(* IEC 61131-3 sources: s7-to-codesys/tests/POUs/ScenariosLang/FB_StarterFbd_ScenarioTest, 10 files *)

(* ---- FB_StarterFbd_ScenarioTest.decl.st ---- *)
// AUTO-GENERATED — не редактировать: s7conv gen-tests, сценарии scenarios/lang/FB_Starter.csv
// Правка — в CSV (scenarios/README.md), затем python -m s7conv build-corpus.
// Назначение: тесты поведения сконвертированного FB_StarterFbd по сценариям CSV (сценариев: 9, строк: 47):
//             один метод-тест на сценарий, строки — по порядку с моделируемым временем GVL_S7Clock.
//             Ожидаемые значения — из CSV (эталонные модели по описанию логики блока), не из
//             результата конвертации.
// Автор:      s7conv 0.1.0 (сгенерировано)
// Версия:     не указана
// Документ:   scenarios/README.md, docs/methodology.md, раздел «Проверка поведения»
FUNCTION_BLOCK FB_StarterFbd_ScenarioTest EXTENDS coUnit.FB_TestSuite
VAR
    fbStartStop : FB_StarterFbd;  // свой экземпляр на сценарий
    xStartStopDone : BOOL;  // сценарий выполнен (выполняется один раз)
    fbStartAndStopTogether : FB_StarterFbd;  // свой экземпляр на сценарий
    xStartAndStopTogetherDone : BOOL;  // сценарий выполнен (выполняется один раз)
    fbInterlockBlocksStart : FB_StarterFbd;  // свой экземпляр на сценарий
    xInterlockBlocksStartDone : BOOL;  // сценарий выполнен (выполняется один раз)
    fbInterlockDropStops : FB_StarterFbd;  // свой экземпляр на сценарий
    xInterlockDropStopsDone : BOOL;  // сценарий выполнен (выполняется один раз)
    fbFeedbackOk : FB_StarterFbd;  // свой экземпляр на сценарий
    xFeedbackOkDone : BOOL;  // сценарий выполнен (выполняется один раз)
    fbFeedbackTimeout : FB_StarterFbd;  // свой экземпляр на сценарий
    xFeedbackTimeoutDone : BOOL;  // сценарий выполнен (выполняется один раз)
    fbFaultResetAndBlock : FB_StarterFbd;  // свой экземпляр на сценарий
    xFaultResetAndBlockDone : BOOL;  // сценарий выполнен (выполняется один раз)
    fbStartCounter : FB_StarterFbd;  // свой экземпляр на сценарий
    xStartCounterDone : BOOL;  // сценарий выполнен (выполняется один раз)
    fbResetWhileRunning : FB_StarterFbd;  // свой экземпляр на сценарий
    xResetWhileRunningDone : BOOL;  // сценарий выполнен (выполняется один раз)
END_VAR

(* ---- FaultResetAndBlock.method.impl.st ---- *)
// AUTO-GENERATED — не редактировать: scenarios/lang/FB_Starter.csv, сценарий FaultResetAndBlock
coUnit.TEST('FaultResetAndBlock');
IF NOT xFaultResetAndBlockDone THEN
    xFaultResetAndBlockDone := TRUE;
    GVL_S7Clock.xSimulation := TRUE;

    // #1, t = 0 мс — Пуск без обратной связи, пуск №1
    GVL_S7Clock.tSimNow := T#0MS;
    fbFaultResetAndBlock.xStart := TRUE;
    fbFaultResetAndBlock.xStop := FALSE;
    fbFaultResetAndBlock.xInterlock := TRUE;
    fbFaultResetAndBlock.xFeedback := FALSE;
    fbFaultResetAndBlock.tFeedbackTime := T#2000MS;
    fbFaultResetAndBlock.xReset := FALSE;
    fbFaultResetAndBlock();
    AssertEquals_BOOL(Expected := TRUE, Actual := fbFaultResetAndBlock.xRun, Message := 'FaultResetAndBlock#1 xRun');
    AssertEquals_BOOL(Expected := FALSE,
                      Actual := fbFaultResetAndBlock.xFault,
                      Message := 'FaultResetAndBlock#1 xFault');
    AssertEquals_INT(Expected := 1, Actual := fbFaultResetAndBlock.iStarts, Message := 'FaultResetAndBlock#1 iStarts');

    // #2, t = 100 мс — ждём
    GVL_S7Clock.tSimNow := T#100MS;
    fbFaultResetAndBlock.xStart := FALSE;
    fbFaultResetAndBlock();
    AssertEquals_BOOL(Expected := TRUE, Actual := fbFaultResetAndBlock.xRun, Message := 'FaultResetAndBlock#2 xRun');
    AssertEquals_BOOL(Expected := FALSE,
                      Actual := fbFaultResetAndBlock.xFault,
                      Message := 'FaultResetAndBlock#2 xFault');
    AssertEquals_INT(Expected := 1, Actual := fbFaultResetAndBlock.iStarts, Message := 'FaultResetAndBlock#2 iStarts');

    // #3, t = 2400 мс — 2.4 с: авария
    GVL_S7Clock.tSimNow := T#2400MS;
    fbFaultResetAndBlock();
    AssertEquals_BOOL(Expected := TRUE, Actual := fbFaultResetAndBlock.xRun, Message := 'FaultResetAndBlock#3 xRun');
    AssertEquals_BOOL(Expected := TRUE,
                      Actual := fbFaultResetAndBlock.xFault,
                      Message := 'FaultResetAndBlock#3 xFault');
    AssertEquals_INT(Expected := 1, Actual := fbFaultResetAndBlock.iStarts, Message := 'FaultResetAndBlock#3 iStarts');

    // #4, t = 2600 мс — Пуск при аварии: R1 = 1 главнее — не включается
    GVL_S7Clock.tSimNow := T#2600MS;
    fbFaultResetAndBlock.xStart := TRUE;
    fbFaultResetAndBlock();
    AssertEquals_BOOL(Expected := FALSE, Actual := fbFaultResetAndBlock.xRun, Message := 'FaultResetAndBlock#4 xRun');
    AssertEquals_BOOL(Expected := TRUE,
                      Actual := fbFaultResetAndBlock.xFault,
                      Message := 'FaultResetAndBlock#4 xFault');
    AssertEquals_INT(Expected := 1, Actual := fbFaultResetAndBlock.iStarts, Message := 'FaultResetAndBlock#4 iStarts');

    // #5, t = 2700 мс — сброс: авария снята
    GVL_S7Clock.tSimNow := T#2700MS;
    fbFaultResetAndBlock.xStart := FALSE;
    fbFaultResetAndBlock.xReset := TRUE;
    fbFaultResetAndBlock();
    AssertEquals_BOOL(Expected := FALSE, Actual := fbFaultResetAndBlock.xRun, Message := 'FaultResetAndBlock#5 xRun');
    AssertEquals_BOOL(Expected := FALSE,
                      Actual := fbFaultResetAndBlock.xFault,
                      Message := 'FaultResetAndBlock#5 xFault');
    AssertEquals_INT(Expected := 1, Actual := fbFaultResetAndBlock.iStarts, Message := 'FaultResetAndBlock#5 iStarts');

    // #6, t = 2800 мс — Пуск: включается, пуск №2
    GVL_S7Clock.tSimNow := T#2800MS;
    fbFaultResetAndBlock.xStart := TRUE;
    fbFaultResetAndBlock.xReset := FALSE;
    fbFaultResetAndBlock();
    AssertEquals_BOOL(Expected := TRUE, Actual := fbFaultResetAndBlock.xRun, Message := 'FaultResetAndBlock#6 xRun');
    AssertEquals_BOOL(Expected := FALSE,
                      Actual := fbFaultResetAndBlock.xFault,
                      Message := 'FaultResetAndBlock#6 xFault');
    AssertEquals_INT(Expected := 2, Actual := fbFaultResetAndBlock.iStarts, Message := 'FaultResetAndBlock#6 iStarts');

    // #7, t = 2900 мс — обратная связь: работает без аварии
    GVL_S7Clock.tSimNow := T#2900MS;
    fbFaultResetAndBlock.xStart := FALSE;
    fbFaultResetAndBlock.xFeedback := TRUE;
    fbFaultResetAndBlock();
    AssertEquals_BOOL(Expected := TRUE, Actual := fbFaultResetAndBlock.xRun, Message := 'FaultResetAndBlock#7 xRun');
    AssertEquals_BOOL(Expected := FALSE,
                      Actual := fbFaultResetAndBlock.xFault,
                      Message := 'FaultResetAndBlock#7 xFault');
    AssertEquals_INT(Expected := 2, Actual := fbFaultResetAndBlock.iStarts, Message := 'FaultResetAndBlock#7 iStarts');

    GVL_S7Clock.xSimulation := FALSE;
END_IF
coUnit.TEST_FINISHED();

(* ---- FeedbackOk.method.impl.st ---- *)
// AUTO-GENERATED — не редактировать: scenarios/lang/FB_Starter.csv, сценарий FeedbackOk
coUnit.TEST('FeedbackOk');
IF NOT xFeedbackOkDone THEN
    xFeedbackOkDone := TRUE;
    GVL_S7Clock.xSimulation := TRUE;

    // #1, t = 0 мс — покой
    GVL_S7Clock.tSimNow := T#0MS;
    fbFeedbackOk.xStart := FALSE;
    fbFeedbackOk.xStop := FALSE;
    fbFeedbackOk.xInterlock := TRUE;
    fbFeedbackOk.xFeedback := FALSE;
    fbFeedbackOk.tFeedbackTime := T#2000MS;
    fbFeedbackOk.xReset := FALSE;
    fbFeedbackOk();
    AssertEquals_BOOL(Expected := FALSE, Actual := fbFeedbackOk.xRun, Message := 'FeedbackOk#1 xRun');
    AssertEquals_BOOL(Expected := FALSE, Actual := fbFeedbackOk.xFault, Message := 'FeedbackOk#1 xFault');
    AssertEquals_INT(Expected := 0, Actual := fbFeedbackOk.iStarts, Message := 'FeedbackOk#1 iStarts');

    // #2, t = 100 мс — Пуск, таймер обратной связи с 0.1 с
    GVL_S7Clock.tSimNow := T#100MS;
    fbFeedbackOk.xStart := TRUE;
    fbFeedbackOk();
    AssertEquals_BOOL(Expected := TRUE, Actual := fbFeedbackOk.xRun, Message := 'FeedbackOk#2 xRun');
    AssertEquals_BOOL(Expected := FALSE, Actual := fbFeedbackOk.xFault, Message := 'FeedbackOk#2 xFault');
    AssertEquals_INT(Expected := 1, Actual := fbFeedbackOk.iStarts, Message := 'FeedbackOk#2 iStarts');

    // #3, t = 1000 мс — обратная связь через 0.9 с
    GVL_S7Clock.tSimNow := T#1000MS;
    fbFeedbackOk.xStart := FALSE;
    fbFeedbackOk.xFeedback := TRUE;
    fbFeedbackOk();
    AssertEquals_BOOL(Expected := TRUE, Actual := fbFeedbackOk.xRun, Message := 'FeedbackOk#3 xRun');
    AssertEquals_BOOL(Expected := FALSE, Actual := fbFeedbackOk.xFault, Message := 'FeedbackOk#3 xFault');
    AssertEquals_INT(Expected := 1, Actual := fbFeedbackOk.iStarts, Message := 'FeedbackOk#3 iStarts');

    // #4, t = 5000 мс — работает, аварии нет
    GVL_S7Clock.tSimNow := T#5000MS;
    fbFeedbackOk();
    AssertEquals_BOOL(Expected := TRUE, Actual := fbFeedbackOk.xRun, Message := 'FeedbackOk#4 xRun');
    AssertEquals_BOOL(Expected := FALSE, Actual := fbFeedbackOk.xFault, Message := 'FeedbackOk#4 xFault');
    AssertEquals_INT(Expected := 1, Actual := fbFeedbackOk.iStarts, Message := 'FeedbackOk#4 iStarts');

    GVL_S7Clock.xSimulation := FALSE;
END_IF
coUnit.TEST_FINISHED();

(* ---- FeedbackTimeout.method.impl.st ---- *)
// AUTO-GENERATED — не редактировать: scenarios/lang/FB_Starter.csv, сценарий FeedbackTimeout
coUnit.TEST('FeedbackTimeout');
IF NOT xFeedbackTimeoutDone THEN
    xFeedbackTimeoutDone := TRUE;
    GVL_S7Clock.xSimulation := TRUE;

    // #1, t = 0 мс — покой
    GVL_S7Clock.tSimNow := T#0MS;
    fbFeedbackTimeout.xStart := FALSE;
    fbFeedbackTimeout.xStop := FALSE;
    fbFeedbackTimeout.xInterlock := TRUE;
    fbFeedbackTimeout.xFeedback := FALSE;
    fbFeedbackTimeout.tFeedbackTime := T#2000MS;
    fbFeedbackTimeout.xReset := FALSE;
    fbFeedbackTimeout();
    AssertEquals_BOOL(Expected := FALSE, Actual := fbFeedbackTimeout.xRun, Message := 'FeedbackTimeout#1 xRun');
    AssertEquals_BOOL(Expected := FALSE, Actual := fbFeedbackTimeout.xFault, Message := 'FeedbackTimeout#1 xFault');
    AssertEquals_INT(Expected := 0, Actual := fbFeedbackTimeout.iStarts, Message := 'FeedbackTimeout#1 iStarts');

    // #2, t = 100 мс — Пуск без обратной связи, таймер с 0.1 с
    GVL_S7Clock.tSimNow := T#100MS;
    fbFeedbackTimeout.xStart := TRUE;
    fbFeedbackTimeout();
    AssertEquals_BOOL(Expected := TRUE, Actual := fbFeedbackTimeout.xRun, Message := 'FeedbackTimeout#2 xRun');
    AssertEquals_BOOL(Expected := FALSE, Actual := fbFeedbackTimeout.xFault, Message := 'FeedbackTimeout#2 xFault');
    AssertEquals_INT(Expected := 1, Actual := fbFeedbackTimeout.iStarts, Message := 'FeedbackTimeout#2 iStarts');

    // #3, t = 1900 мс — 1.8 с < 2 с: аварии нет
    GVL_S7Clock.tSimNow := T#1900MS;
    fbFeedbackTimeout.xStart := FALSE;
    fbFeedbackTimeout();
    AssertEquals_BOOL(Expected := TRUE, Actual := fbFeedbackTimeout.xRun, Message := 'FeedbackTimeout#3 xRun');
    AssertEquals_BOOL(Expected := FALSE, Actual := fbFeedbackTimeout.xFault, Message := 'FeedbackTimeout#3 xFault');
    AssertEquals_INT(Expected := 1, Actual := fbFeedbackTimeout.iStarts, Message := 'FeedbackTimeout#3 iStarts');

    // #4, t = 2100 мс, на пороге таймера — 2.0 с = tFeedbackTime: авария; xRun ещё TRUE (сеть 1 раньше сети 3)
    GVL_S7Clock.tSimNow := T#2100MS;
    fbFeedbackTimeout();
    AssertEquals_BOOL(Expected := TRUE, Actual := fbFeedbackTimeout.xRun, Message := 'FeedbackTimeout#4 xRun');
    AssertEquals_BOOL(Expected := TRUE, Actual := fbFeedbackTimeout.xFault, Message := 'FeedbackTimeout#4 xFault');
    AssertEquals_INT(Expected := 1, Actual := fbFeedbackTimeout.iStarts, Message := 'FeedbackTimeout#4 iStarts');

    // #5, t = 2300 мс — R1 = xFault: насос выключен, авария держится
    GVL_S7Clock.tSimNow := T#2300MS;
    fbFeedbackTimeout();
    AssertEquals_BOOL(Expected := FALSE, Actual := fbFeedbackTimeout.xRun, Message := 'FeedbackTimeout#5 xRun');
    AssertEquals_BOOL(Expected := TRUE, Actual := fbFeedbackTimeout.xFault, Message := 'FeedbackTimeout#5 xFault');
    AssertEquals_INT(Expected := 1, Actual := fbFeedbackTimeout.iStarts, Message := 'FeedbackTimeout#5 iStarts');

    // #6, t = 3000 мс — авария держится (самоподхват)
    GVL_S7Clock.tSimNow := T#3000MS;
    fbFeedbackTimeout();
    AssertEquals_BOOL(Expected := FALSE, Actual := fbFeedbackTimeout.xRun, Message := 'FeedbackTimeout#6 xRun');
    AssertEquals_BOOL(Expected := TRUE, Actual := fbFeedbackTimeout.xFault, Message := 'FeedbackTimeout#6 xFault');
    AssertEquals_INT(Expected := 1, Actual := fbFeedbackTimeout.iStarts, Message := 'FeedbackTimeout#6 iStarts');

    GVL_S7Clock.xSimulation := FALSE;
END_IF
coUnit.TEST_FINISHED();

(* ---- InterlockBlocksStart.method.impl.st ---- *)
// AUTO-GENERATED — не редактировать: scenarios/lang/FB_Starter.csv, сценарий InterlockBlocksStart
coUnit.TEST('InterlockBlocksStart');
IF NOT xInterlockBlocksStartDone THEN
    xInterlockBlocksStartDone := TRUE;
    GVL_S7Clock.xSimulation := TRUE;

    // #1, t = 0 мс — блокировка
    GVL_S7Clock.tSimNow := T#0MS;
    fbInterlockBlocksStart.xStart := FALSE;
    fbInterlockBlocksStart.xStop := FALSE;
    fbInterlockBlocksStart.xInterlock := FALSE;
    fbInterlockBlocksStart.xFeedback := FALSE;
    fbInterlockBlocksStart.tFeedbackTime := T#2000MS;
    fbInterlockBlocksStart.xReset := FALSE;
    fbInterlockBlocksStart();
    AssertEquals_BOOL(Expected := FALSE,
                      Actual := fbInterlockBlocksStart.xRun,
                      Message := 'InterlockBlocksStart#1 xRun');
    AssertEquals_BOOL(Expected := FALSE,
                      Actual := fbInterlockBlocksStart.xFault,
                      Message := 'InterlockBlocksStart#1 xFault');
    AssertEquals_INT(Expected := 0,
                     Actual := fbInterlockBlocksStart.iStarts,
                     Message := 'InterlockBlocksStart#1 iStarts');

    // #2, t = 100 мс — Пуск при блокировке: не включается
    GVL_S7Clock.tSimNow := T#100MS;
    fbInterlockBlocksStart.xStart := TRUE;
    fbInterlockBlocksStart();
    AssertEquals_BOOL(Expected := FALSE,
                      Actual := fbInterlockBlocksStart.xRun,
                      Message := 'InterlockBlocksStart#2 xRun');
    AssertEquals_BOOL(Expected := FALSE,
                      Actual := fbInterlockBlocksStart.xFault,
                      Message := 'InterlockBlocksStart#2 xFault');
    AssertEquals_INT(Expected := 0,
                     Actual := fbInterlockBlocksStart.iStarts,
                     Message := 'InterlockBlocksStart#2 iStarts');

    // #3, t = 200 мс — кнопка отпущена
    GVL_S7Clock.tSimNow := T#200MS;
    fbInterlockBlocksStart.xStart := FALSE;
    fbInterlockBlocksStart();
    AssertEquals_BOOL(Expected := FALSE,
                      Actual := fbInterlockBlocksStart.xRun,
                      Message := 'InterlockBlocksStart#3 xRun');
    AssertEquals_BOOL(Expected := FALSE,
                      Actual := fbInterlockBlocksStart.xFault,
                      Message := 'InterlockBlocksStart#3 xFault');
    AssertEquals_INT(Expected := 0,
                     Actual := fbInterlockBlocksStart.iStarts,
                     Message := 'InterlockBlocksStart#3 iStarts');

    // #4, t = 300 мс — блокировка снята: пуск не запомнен
    GVL_S7Clock.tSimNow := T#300MS;
    fbInterlockBlocksStart.xInterlock := TRUE;
    fbInterlockBlocksStart();
    AssertEquals_BOOL(Expected := FALSE,
                      Actual := fbInterlockBlocksStart.xRun,
                      Message := 'InterlockBlocksStart#4 xRun');
    AssertEquals_BOOL(Expected := FALSE,
                      Actual := fbInterlockBlocksStart.xFault,
                      Message := 'InterlockBlocksStart#4 xFault');
    AssertEquals_INT(Expected := 0,
                     Actual := fbInterlockBlocksStart.iStarts,
                     Message := 'InterlockBlocksStart#4 iStarts');

    // #5, t = 400 мс — новый Пуск: включается, пуск №1
    GVL_S7Clock.tSimNow := T#400MS;
    fbInterlockBlocksStart.xStart := TRUE;
    fbInterlockBlocksStart();
    AssertEquals_BOOL(Expected := TRUE,
                      Actual := fbInterlockBlocksStart.xRun,
                      Message := 'InterlockBlocksStart#5 xRun');
    AssertEquals_BOOL(Expected := FALSE,
                      Actual := fbInterlockBlocksStart.xFault,
                      Message := 'InterlockBlocksStart#5 xFault');
    AssertEquals_INT(Expected := 1,
                     Actual := fbInterlockBlocksStart.iStarts,
                     Message := 'InterlockBlocksStart#5 iStarts');

    GVL_S7Clock.xSimulation := FALSE;
END_IF
coUnit.TEST_FINISHED();

(* ---- InterlockDropStops.method.impl.st ---- *)
// AUTO-GENERATED — не редактировать: scenarios/lang/FB_Starter.csv, сценарий InterlockDropStops
coUnit.TEST('InterlockDropStops');
IF NOT xInterlockDropStopsDone THEN
    xInterlockDropStopsDone := TRUE;
    GVL_S7Clock.xSimulation := TRUE;

    // #1, t = 0 мс — Пуск, пуск №1
    GVL_S7Clock.tSimNow := T#0MS;
    fbInterlockDropStops.xStart := TRUE;
    fbInterlockDropStops.xStop := FALSE;
    fbInterlockDropStops.xInterlock := TRUE;
    fbInterlockDropStops.xFeedback := FALSE;
    fbInterlockDropStops.tFeedbackTime := T#2000MS;
    fbInterlockDropStops.xReset := FALSE;
    fbInterlockDropStops();
    AssertEquals_BOOL(Expected := TRUE, Actual := fbInterlockDropStops.xRun, Message := 'InterlockDropStops#1 xRun');
    AssertEquals_BOOL(Expected := FALSE,
                      Actual := fbInterlockDropStops.xFault,
                      Message := 'InterlockDropStops#1 xFault');
    AssertEquals_INT(Expected := 1, Actual := fbInterlockDropStops.iStarts, Message := 'InterlockDropStops#1 iStarts');

    // #2, t = 100 мс — работает
    GVL_S7Clock.tSimNow := T#100MS;
    fbInterlockDropStops.xStart := FALSE;
    fbInterlockDropStops.xFeedback := TRUE;
    fbInterlockDropStops();
    AssertEquals_BOOL(Expected := TRUE, Actual := fbInterlockDropStops.xRun, Message := 'InterlockDropStops#2 xRun');
    AssertEquals_BOOL(Expected := FALSE,
                      Actual := fbInterlockDropStops.xFault,
                      Message := 'InterlockDropStops#2 xFault');
    AssertEquals_INT(Expected := 1, Actual := fbInterlockDropStops.iStarts, Message := 'InterlockDropStops#2 iStarts');

    // #3, t = 500 мс — блокировка пропала: выключается
    GVL_S7Clock.tSimNow := T#500MS;
    fbInterlockDropStops.xInterlock := FALSE;
    fbInterlockDropStops();
    AssertEquals_BOOL(Expected := FALSE, Actual := fbInterlockDropStops.xRun, Message := 'InterlockDropStops#3 xRun');
    AssertEquals_BOOL(Expected := FALSE,
                      Actual := fbInterlockDropStops.xFault,
                      Message := 'InterlockDropStops#3 xFault');
    AssertEquals_INT(Expected := 1, Actual := fbInterlockDropStops.iStarts, Message := 'InterlockDropStops#3 iStarts');

    // #4, t = 600 мс — блокировка вернулась: остаётся выключенным
    GVL_S7Clock.tSimNow := T#600MS;
    fbInterlockDropStops.xInterlock := TRUE;
    fbInterlockDropStops.xFeedback := FALSE;
    fbInterlockDropStops();
    AssertEquals_BOOL(Expected := FALSE, Actual := fbInterlockDropStops.xRun, Message := 'InterlockDropStops#4 xRun');
    AssertEquals_BOOL(Expected := FALSE,
                      Actual := fbInterlockDropStops.xFault,
                      Message := 'InterlockDropStops#4 xFault');
    AssertEquals_INT(Expected := 1, Actual := fbInterlockDropStops.iStarts, Message := 'InterlockDropStops#4 iStarts');

    GVL_S7Clock.xSimulation := FALSE;
END_IF
coUnit.TEST_FINISHED();

(* ---- ResetWhileRunning.method.impl.st ---- *)
// AUTO-GENERATED — не редактировать: scenarios/lang/FB_Starter.csv, сценарий ResetWhileRunning
coUnit.TEST('ResetWhileRunning');
IF NOT xResetWhileRunningDone THEN
    xResetWhileRunningDone := TRUE;
    GVL_S7Clock.xSimulation := TRUE;

    // #1, t = 0 мс — пуск №1
    GVL_S7Clock.tSimNow := T#0MS;
    fbResetWhileRunning.xStart := TRUE;
    fbResetWhileRunning.xStop := FALSE;
    fbResetWhileRunning.xInterlock := TRUE;
    fbResetWhileRunning.xFeedback := TRUE;
    fbResetWhileRunning.tFeedbackTime := T#2000MS;
    fbResetWhileRunning.xReset := FALSE;
    fbResetWhileRunning();
    AssertEquals_BOOL(Expected := TRUE, Actual := fbResetWhileRunning.xRun, Message := 'ResetWhileRunning#1 xRun');
    AssertEquals_BOOL(Expected := FALSE, Actual := fbResetWhileRunning.xFault, Message := 'ResetWhileRunning#1 xFault');
    AssertEquals_INT(Expected := 1, Actual := fbResetWhileRunning.iStarts, Message := 'ResetWhileRunning#1 iStarts');

    // #2, t = 100 мс — сброс в работе: без изменений
    GVL_S7Clock.tSimNow := T#100MS;
    fbResetWhileRunning.xStart := FALSE;
    fbResetWhileRunning.xReset := TRUE;
    fbResetWhileRunning();
    AssertEquals_BOOL(Expected := TRUE, Actual := fbResetWhileRunning.xRun, Message := 'ResetWhileRunning#2 xRun');
    AssertEquals_BOOL(Expected := FALSE, Actual := fbResetWhileRunning.xFault, Message := 'ResetWhileRunning#2 xFault');
    AssertEquals_INT(Expected := 1, Actual := fbResetWhileRunning.iStarts, Message := 'ResetWhileRunning#2 iStarts');

    // #3, t = 200 мс — Пуск в работе: SR уже установлен, счёта нет
    GVL_S7Clock.tSimNow := T#200MS;
    fbResetWhileRunning.xStart := TRUE;
    fbResetWhileRunning.xReset := FALSE;
    fbResetWhileRunning();
    AssertEquals_BOOL(Expected := TRUE, Actual := fbResetWhileRunning.xRun, Message := 'ResetWhileRunning#3 xRun');
    AssertEquals_BOOL(Expected := FALSE, Actual := fbResetWhileRunning.xFault, Message := 'ResetWhileRunning#3 xFault');
    AssertEquals_INT(Expected := 1, Actual := fbResetWhileRunning.iStarts, Message := 'ResetWhileRunning#3 iStarts');

    // #4, t = 300 мс — работает
    GVL_S7Clock.tSimNow := T#300MS;
    fbResetWhileRunning.xStart := FALSE;
    fbResetWhileRunning();
    AssertEquals_BOOL(Expected := TRUE, Actual := fbResetWhileRunning.xRun, Message := 'ResetWhileRunning#4 xRun');
    AssertEquals_BOOL(Expected := FALSE, Actual := fbResetWhileRunning.xFault, Message := 'ResetWhileRunning#4 xFault');
    AssertEquals_INT(Expected := 1, Actual := fbResetWhileRunning.iStarts, Message := 'ResetWhileRunning#4 iStarts');

    GVL_S7Clock.xSimulation := FALSE;
END_IF
coUnit.TEST_FINISHED();

(* ---- StartAndStopTogether.method.impl.st ---- *)
// AUTO-GENERATED — не редактировать: scenarios/lang/FB_Starter.csv, сценарий StartAndStopTogether
coUnit.TEST('StartAndStopTogether');
IF NOT xStartAndStopTogetherDone THEN
    xStartAndStopTogetherDone := TRUE;
    GVL_S7Clock.xSimulation := TRUE;

    // #1, t = 0 мс — покой
    GVL_S7Clock.tSimNow := T#0MS;
    fbStartAndStopTogether.xStart := FALSE;
    fbStartAndStopTogether.xStop := FALSE;
    fbStartAndStopTogether.xInterlock := TRUE;
    fbStartAndStopTogether.xFeedback := FALSE;
    fbStartAndStopTogether.tFeedbackTime := T#2000MS;
    fbStartAndStopTogether.xReset := FALSE;
    fbStartAndStopTogether();
    AssertEquals_BOOL(Expected := FALSE,
                      Actual := fbStartAndStopTogether.xRun,
                      Message := 'StartAndStopTogether#1 xRun');
    AssertEquals_BOOL(Expected := FALSE,
                      Actual := fbStartAndStopTogether.xFault,
                      Message := 'StartAndStopTogether#1 xFault');
    AssertEquals_INT(Expected := 0,
                     Actual := fbStartAndStopTogether.iStarts,
                     Message := 'StartAndStopTogether#1 iStarts');

    // #2, t = 100 мс — S = R1 = 1: не включается
    GVL_S7Clock.tSimNow := T#100MS;
    fbStartAndStopTogether.xStart := TRUE;
    fbStartAndStopTogether.xStop := TRUE;
    fbStartAndStopTogether();
    AssertEquals_BOOL(Expected := FALSE,
                      Actual := fbStartAndStopTogether.xRun,
                      Message := 'StartAndStopTogether#2 xRun');
    AssertEquals_BOOL(Expected := FALSE,
                      Actual := fbStartAndStopTogether.xFault,
                      Message := 'StartAndStopTogether#2 xFault');
    AssertEquals_INT(Expected := 0,
                     Actual := fbStartAndStopTogether.iStarts,
                     Message := 'StartAndStopTogether#2 iStarts');

    // #3, t = 200 мс — Стоп отпущен, Пуск держится: включается, пуск №1
    GVL_S7Clock.tSimNow := T#200MS;
    fbStartAndStopTogether.xStop := FALSE;
    fbStartAndStopTogether();
    AssertEquals_BOOL(Expected := TRUE,
                      Actual := fbStartAndStopTogether.xRun,
                      Message := 'StartAndStopTogether#3 xRun');
    AssertEquals_BOOL(Expected := FALSE,
                      Actual := fbStartAndStopTogether.xFault,
                      Message := 'StartAndStopTogether#3 xFault');
    AssertEquals_INT(Expected := 1,
                     Actual := fbStartAndStopTogether.iStarts,
                     Message := 'StartAndStopTogether#3 iStarts');

    // #4, t = 300 мс — работает
    GVL_S7Clock.tSimNow := T#300MS;
    fbStartAndStopTogether.xStart := FALSE;
    fbStartAndStopTogether.xFeedback := TRUE;
    fbStartAndStopTogether();
    AssertEquals_BOOL(Expected := TRUE,
                      Actual := fbStartAndStopTogether.xRun,
                      Message := 'StartAndStopTogether#4 xRun');
    AssertEquals_BOOL(Expected := FALSE,
                      Actual := fbStartAndStopTogether.xFault,
                      Message := 'StartAndStopTogether#4 xFault');
    AssertEquals_INT(Expected := 1,
                     Actual := fbStartAndStopTogether.iStarts,
                     Message := 'StartAndStopTogether#4 iStarts');

    // #5, t = 400 мс — в работе снова S = R1 = 1: выключается
    GVL_S7Clock.tSimNow := T#400MS;
    fbStartAndStopTogether.xStart := TRUE;
    fbStartAndStopTogether.xStop := TRUE;
    fbStartAndStopTogether();
    AssertEquals_BOOL(Expected := FALSE,
                      Actual := fbStartAndStopTogether.xRun,
                      Message := 'StartAndStopTogether#5 xRun');
    AssertEquals_BOOL(Expected := FALSE,
                      Actual := fbStartAndStopTogether.xFault,
                      Message := 'StartAndStopTogether#5 xFault');
    AssertEquals_INT(Expected := 1,
                     Actual := fbStartAndStopTogether.iStarts,
                     Message := 'StartAndStopTogether#5 iStarts');

    // #6, t = 500 мс — выключен
    GVL_S7Clock.tSimNow := T#500MS;
    fbStartAndStopTogether.xStart := FALSE;
    fbStartAndStopTogether.xStop := FALSE;
    fbStartAndStopTogether.xFeedback := FALSE;
    fbStartAndStopTogether();
    AssertEquals_BOOL(Expected := FALSE,
                      Actual := fbStartAndStopTogether.xRun,
                      Message := 'StartAndStopTogether#6 xRun');
    AssertEquals_BOOL(Expected := FALSE,
                      Actual := fbStartAndStopTogether.xFault,
                      Message := 'StartAndStopTogether#6 xFault');
    AssertEquals_INT(Expected := 1,
                     Actual := fbStartAndStopTogether.iStarts,
                     Message := 'StartAndStopTogether#6 iStarts');

    GVL_S7Clock.xSimulation := FALSE;
END_IF
coUnit.TEST_FINISHED();

(* ---- StartCounter.method.impl.st ---- *)
// AUTO-GENERATED — не редактировать: scenarios/lang/FB_Starter.csv, сценарий StartCounter
coUnit.TEST('StartCounter');
IF NOT xStartCounterDone THEN
    xStartCounterDone := TRUE;
    GVL_S7Clock.xSimulation := TRUE;

    // #1, t = 0 мс — пуск №1
    GVL_S7Clock.tSimNow := T#0MS;
    fbStartCounter.xStart := TRUE;
    fbStartCounter.xStop := FALSE;
    fbStartCounter.xInterlock := TRUE;
    fbStartCounter.xFeedback := TRUE;
    fbStartCounter.tFeedbackTime := T#2000MS;
    fbStartCounter.xReset := FALSE;
    fbStartCounter();
    AssertEquals_BOOL(Expected := TRUE, Actual := fbStartCounter.xRun, Message := 'StartCounter#1 xRun');
    AssertEquals_BOOL(Expected := FALSE, Actual := fbStartCounter.xFault, Message := 'StartCounter#1 xFault');
    AssertEquals_INT(Expected := 1, Actual := fbStartCounter.iStarts, Message := 'StartCounter#1 iStarts');

    // #2, t = 100 мс — Пуск держится: без нового счёта
    GVL_S7Clock.tSimNow := T#100MS;
    fbStartCounter();
    AssertEquals_BOOL(Expected := TRUE, Actual := fbStartCounter.xRun, Message := 'StartCounter#2 xRun');
    AssertEquals_BOOL(Expected := FALSE, Actual := fbStartCounter.xFault, Message := 'StartCounter#2 xFault');
    AssertEquals_INT(Expected := 1, Actual := fbStartCounter.iStarts, Message := 'StartCounter#2 iStarts');

    // #3, t = 200 мс — стоп
    GVL_S7Clock.tSimNow := T#200MS;
    fbStartCounter.xStart := FALSE;
    fbStartCounter.xStop := TRUE;
    fbStartCounter();
    AssertEquals_BOOL(Expected := FALSE, Actual := fbStartCounter.xRun, Message := 'StartCounter#3 xRun');
    AssertEquals_BOOL(Expected := FALSE, Actual := fbStartCounter.xFault, Message := 'StartCounter#3 xFault');
    AssertEquals_INT(Expected := 1, Actual := fbStartCounter.iStarts, Message := 'StartCounter#3 iStarts');

    // #4, t = 300 мс — пуск №2
    GVL_S7Clock.tSimNow := T#300MS;
    fbStartCounter.xStart := TRUE;
    fbStartCounter.xStop := FALSE;
    fbStartCounter();
    AssertEquals_BOOL(Expected := TRUE, Actual := fbStartCounter.xRun, Message := 'StartCounter#4 xRun');
    AssertEquals_BOOL(Expected := FALSE, Actual := fbStartCounter.xFault, Message := 'StartCounter#4 xFault');
    AssertEquals_INT(Expected := 2, Actual := fbStartCounter.iStarts, Message := 'StartCounter#4 iStarts');

    // #5, t = 400 мс — стоп
    GVL_S7Clock.tSimNow := T#400MS;
    fbStartCounter.xStart := FALSE;
    fbStartCounter.xStop := TRUE;
    fbStartCounter();
    AssertEquals_BOOL(Expected := FALSE, Actual := fbStartCounter.xRun, Message := 'StartCounter#5 xRun');
    AssertEquals_BOOL(Expected := FALSE, Actual := fbStartCounter.xFault, Message := 'StartCounter#5 xFault');
    AssertEquals_INT(Expected := 2, Actual := fbStartCounter.iStarts, Message := 'StartCounter#5 iStarts');

    // #6, t = 500 мс — покой: 2 пуска
    GVL_S7Clock.tSimNow := T#500MS;
    fbStartCounter.xStop := FALSE;
    fbStartCounter();
    AssertEquals_BOOL(Expected := FALSE, Actual := fbStartCounter.xRun, Message := 'StartCounter#6 xRun');
    AssertEquals_BOOL(Expected := FALSE, Actual := fbStartCounter.xFault, Message := 'StartCounter#6 xFault');
    AssertEquals_INT(Expected := 2, Actual := fbStartCounter.iStarts, Message := 'StartCounter#6 iStarts');

    GVL_S7Clock.xSimulation := FALSE;
END_IF
coUnit.TEST_FINISHED();

(* ---- StartStop.method.impl.st ---- *)
// AUTO-GENERATED — не редактировать: scenarios/lang/FB_Starter.csv, сценарий StartStop
coUnit.TEST('StartStop');
IF NOT xStartStopDone THEN
    xStartStopDone := TRUE;
    GVL_S7Clock.xSimulation := TRUE;

    // #1, t = 0 мс — покой
    GVL_S7Clock.tSimNow := T#0MS;
    fbStartStop.xStart := FALSE;
    fbStartStop.xStop := FALSE;
    fbStartStop.xInterlock := TRUE;
    fbStartStop.xFeedback := FALSE;
    fbStartStop.tFeedbackTime := T#2000MS;
    fbStartStop.xReset := FALSE;
    fbStartStop();
    AssertEquals_BOOL(Expected := FALSE, Actual := fbStartStop.xRun, Message := 'StartStop#1 xRun');
    AssertEquals_BOOL(Expected := FALSE, Actual := fbStartStop.xFault, Message := 'StartStop#1 xFault');
    AssertEquals_INT(Expected := 0, Actual := fbStartStop.iStarts, Message := 'StartStop#1 iStarts');

    // #2, t = 100 мс — Пуск: SR установлен, пуск №1
    GVL_S7Clock.tSimNow := T#100MS;
    fbStartStop.xStart := TRUE;
    fbStartStop();
    AssertEquals_BOOL(Expected := TRUE, Actual := fbStartStop.xRun, Message := 'StartStop#2 xRun');
    AssertEquals_BOOL(Expected := FALSE, Actual := fbStartStop.xFault, Message := 'StartStop#2 xFault');
    AssertEquals_INT(Expected := 1, Actual := fbStartStop.iStarts, Message := 'StartStop#2 iStarts');

    // #3, t = 200 мс — кнопка отпущена, обратная связь: работает
    GVL_S7Clock.tSimNow := T#200MS;
    fbStartStop.xStart := FALSE;
    fbStartStop.xFeedback := TRUE;
    fbStartStop();
    AssertEquals_BOOL(Expected := TRUE, Actual := fbStartStop.xRun, Message := 'StartStop#3 xRun');
    AssertEquals_BOOL(Expected := FALSE, Actual := fbStartStop.xFault, Message := 'StartStop#3 xFault');
    AssertEquals_INT(Expected := 1, Actual := fbStartStop.iStarts, Message := 'StartStop#3 iStarts');

    // #4, t = 1000 мс — Стоп: SR сброшен
    GVL_S7Clock.tSimNow := T#1000MS;
    fbStartStop.xStop := TRUE;
    fbStartStop();
    AssertEquals_BOOL(Expected := FALSE, Actual := fbStartStop.xRun, Message := 'StartStop#4 xRun');
    AssertEquals_BOOL(Expected := FALSE, Actual := fbStartStop.xFault, Message := 'StartStop#4 xFault');
    AssertEquals_INT(Expected := 1, Actual := fbStartStop.iStarts, Message := 'StartStop#4 iStarts');

    // #5, t = 1100 мс — стоп отпущен: остаётся выключенным
    GVL_S7Clock.tSimNow := T#1100MS;
    fbStartStop.xStop := FALSE;
    fbStartStop.xFeedback := FALSE;
    fbStartStop();
    AssertEquals_BOOL(Expected := FALSE, Actual := fbStartStop.xRun, Message := 'StartStop#5 xRun');
    AssertEquals_BOOL(Expected := FALSE, Actual := fbStartStop.xFault, Message := 'StartStop#5 xFault');
    AssertEquals_INT(Expected := 1, Actual := fbStartStop.iStarts, Message := 'StartStop#5 iStarts');

    GVL_S7Clock.xSimulation := FALSE;
END_IF
coUnit.TEST_FINISHED();
